(* IEC 61131-3 sources: plc-process-lib/tests/POUs/Helpers/FB_TestDeviceExt, 2 files *)

(* ---- FB_TestDeviceExt.decl.st ---- *)
// Назначение: наследник второго уровня FB_TestDevice для проверок времени выполнения R2 и R3
//             контракта: тело вызывает тело FB_TestDevice через SUPER^ со всеми VAR_IN_OUT,
//             до вызова пишет точку расширения, после — унаследованный stCmd; хук OnModeChanged
//             переопределён ещё раз (виртуальный вызов THIS^ из метода базы). Только для тестов.
// Автор:      kr0nsch
// Версия:     0.1.0
// Документ:   docs/TESTING.md, раздел «Тестовое устройство»
FUNCTION_BLOCK FB_TestDeviceExt EXTENDS FB_TestDevice
VAR_INPUT
    xExtFault : BOOL;            // доп. причина отказа — в точку расширения xFaultAdd до SUPER^
END_VAR
VAR
    uiExtBodyCalls : UINT;       // сколько раз выполнено это тело
    uiExtHookCalls : UINT;       // вызовов этой части хука
END_VAR

(* ---- OnModeChanged.method.decl.st ---- *)
// Хук второго уровня: сначала FB_TestDevice (SUPER^), затем своя часть (цифра 2 в udiHookTrace)
METHOD PROTECTED OnModeChanged
VAR_INPUT
    eOld : E_DeviceMode;   // режим до смены
    eNew : E_DeviceMode;   // новый режим
END_VAR
